(* IEC 61131-3 sources: SHRDCAssessment/openplc, 1 file *)

(* ---- tracer_bullet.st ---- *)
PROGRAM TracerBullet
  VAR
    PhotoEye AT %IX0.4 : BOOL;
    Conveyor_Run AT %QX0.0 : BOOL;
  END_VAR

  Conveyor_Run := NOT PhotoEye;
END_PROGRAM

CONFIGURATION Config0
  RESOURCE Res0 ON PLC
    TASK task0(INTERVAL := T#20ms, PRIORITY := 0);
    PROGRAM instance0 WITH task0 : TracerBullet;
  END_RESOURCE
END_CONFIGURATION
